Staubli VAL3: moveJToJoint.pgx

public program moveJToJoint(joint x_jTarget, tool x_tTool, mdesc x_mSpeed)
// //作用：用关节运动的方式移动到目标点。
//   //参数：
//   //x_jTarget: 目标点Joint值
//   //  x_tTool：去目标点使用的工具值
//   //  x_mSpeed:去目标点使用的速度值
//   //x_bWaitEndmove:到达目标点，没有混合，为true则是严格到达目标点
  local bool l_bInRange
begin
  //作用：用关节运动的方式移动到目标点。
  //参数：
  //x_jTarget: 目标点Joint值
  //  x_tTool：去目标点使用的工具值
  //  x_mSpeed:去目标点使用的速度值
  //  x_bWaitEndmove:到达目标点，没有混合，为true则是严格到达目标点

  l_bInRange=isInRange(x_jTarget)
  if l_bInRange==true
    nMoveIDRef=movej(x_jTarget,x_tTool,x_mSpeed)
    call checkMoveId()
  else
    //超出机器人限位
    call rs:setAlarm(221,-1)
  endIf

end
